Fanuc KAREL source: KO00002.KL

PROGRAM KO00002
%NOLOCKGROUP
VAR
  P1: POSITION
  P2: POSITION
  P3: POSITION
  OUT: XYZWPR
BEGIN
  OUT = FRAME(P1, P2, P3)
END KO00002
